(* IEC 61131-3 sources: codesys-elevator/codesys/src, 10 files *)

(* ---- E_Direction.st ---- *)
(* ==========================================================================
   E_Direction : かごの進行方向（Modbus の IR3 にそのまま載る）
   ========================================================================== *)
{attribute 'qualified_only'}   (* CODESYS 独自: E_Direction.Up の形でしか書けないようにする *)
TYPE E_Direction :
(
    Stop := 0,
    Up   := 1,
    Down := 2
) INT;
END_TYPE

(* ---- E_ElevCmd.st ---- *)
(* ==========================================================================
   E_ElevCmd : 画面から送られてくる指令の種類（Modbus の HR0 の値）
   ========================================================================== *)
{attribute 'qualified_only'}   (* CODESYS 独自: E_ElevCmd.CarCall の形でしか書けないようにする *)
TYPE E_ElevCmd :
(
    None      := 0,
    CarCall   := 1,   (* かご内の行き先ボタン（対象階 = HR1） *)
    HallCall  := 2,   (* 乗り場の呼びボタン（対象階 = HR1） *)
    DoorOpen  := 3,   (* 「開」ボタン *)
    DoorClose := 4    (* 「閉」ボタン *)
) INT;
END_TYPE

(* ---- E_ElevState.st ---- *)
(* ==========================================================================
   E_ElevState : エレベータの状態
   値は Modbus の IR0 にそのまま載り、画面（web/src/config.ts）と対応しているので、
   番号を変えないこと
   ========================================================================== *)
{attribute 'qualified_only'}   (* CODESYS 独自: E_ElevState.Idle の形でしか書けないようにする *)
TYPE E_ElevState :
(
    Idle        := 0,   (* 扉を閉めて停止中 *)
    DoorOpening := 1,   (* 扉を開けている途中 *)
    DoorOpen    := 2,   (* 扉が開いている（乗り降り中） *)
    DoorClosing := 3,   (* 扉を閉めている途中 *)
    Moving      := 4,   (* 移動中 *)
    Overload    := 5    (* 重量・人数オーバー。扉を開けたまま警報 *)
) INT;
END_TYPE

(* ---- GVL_ElevIO.st ---- *)
(* ==========================================================================
   GVL_ElevIO : Modbus TCP Slave の I/O マッピング先
   ・aElevToTS   → ModbusTCP Slave の「Input Registers」(%QW) にマッピング（20 個）
   ・aElevFromTS → ModbusTCP Slave の「Holding Registers」(%IW) にマッピング（10 個）
   各レジスタの意味は README.md のレジスタマップ表を参照
   ========================================================================== *)
{attribute 'qualified_only'}   (* CODESYS 独自: GVL_ElevIO.aElevToTS の形でしか書けないようにする *)
VAR_GLOBAL
    aElevToTS   : ARRAY[0..19] OF WORD;   (* PLC → TypeScript（FC04 で読まれる） *)
    aElevFromTS : ARRAY[0..9]  OF WORD;   (* TypeScript → PLC（FC16 で書かれる） *)
END_VAR

(* ---- GVL_ElevParam.st ---- *)
(* ==========================================================================
   GVL_ElevParam : エレベータの仕様（定数）
   画面側（web/src/config.ts）は IR11〜13 で受け取った値を使うので、
   ここを変えれば画面も追従する（FLOOR_COUNT は最大 16）
   ========================================================================== *)
{attribute 'qualified_only'}   (* CODESYS 独自: GVL_ElevParam.FLOOR_COUNT の形でしか書けないようにする *)
VAR_GLOBAL CONSTANT
    FLOOR_COUNT        : INT  := 5;       (* 階数 [階]。1F〜5F。呼びは WORD のビットで持つので最大 16 *)
    MAX_LOAD_KG        : INT  := 600;     (* 定格積載量 [kg] *)
    MAX_PERSONS        : INT  := 9;       (* 定員 [人] *)
    SPEED_FLOORS_PER_S : REAL := 0.5;     (* かごの速さ [階/s] *)
    DOOR_TRAVEL        : TIME := T#2S;    (* 扉が全閉から全開になるまでの時間 *)
    DOOR_DWELL         : TIME := T#5S;    (* 扉を開けておく時間（閉ボタンで短縮できる） *)
    POSITION_EPS       : REAL := 0.001;   (* 階に着いたかの判定の許容差 [階] *)
END_VAR

(* ---- FC_FloorBit.st ---- *)
(* ==========================================================================
   FC_FloorBit
   目的 : 階番号を、呼びを表す WORD のビットに変換する（bit0 = 1F）
   入力 : nFloor  階 [1..FLOOR_COUNT]
   戻り : 該当ビットだけ立った WORD。範囲外の階は 0（呼びとして扱わない）
   履歴 : 2026-10-19  初版
   ========================================================================== *)
FUNCTION FC_FloorBit : WORD
VAR_INPUT
    nFloor : INT;
END_VAR

IF nFloor >= 1 AND nFloor <= GVL_ElevParam.FLOOR_COUNT THEN
    FC_FloorBit := SHL(WORD#1, nFloor - 1);
ELSE
    FC_FloorBit := 0;   (* 画面から範囲外の階が来ても、存在しない階を呼ばない *)
END_IF

(* ---- FC_NextCallFloor.st ---- *)
(* ==========================================================================
   FC_NextCallFloor
   目的 : 進行方向の先にある、いちばん近い呼びの階を探す
          （エレベータの基本的な運転方式：今の方向の呼びを順に片付けてから折り返す）
   入力 : wCalls      呼び（かご内 OR 乗り場。bit0 = 1F）
          rPosition   かごの現在位置 [階]
          eDirection  探す方向
   戻り : 見つかった階 [1..FLOOR_COUNT]。無ければ 0
   履歴 : 2026-10-19  初版
   ========================================================================== *)
FUNCTION FC_NextCallFloor : INT
VAR_INPUT
    wCalls     : WORD;
    rPosition  : REAL;
    eDirection : E_Direction;
END_VAR
VAR
    nFloor : INT;
END_VAR

FC_NextCallFloor := 0;

CASE eDirection OF
    E_Direction.Up:
        (* 下から順に見て、今の位置以上で最初に見つかった呼び *)
        FOR nFloor := 1 TO GVL_ElevParam.FLOOR_COUNT DO
            IF (wCalls AND FC_FloorBit(nFloor)) <> 0
               AND INT_TO_REAL(nFloor) >= rPosition - GVL_ElevParam.POSITION_EPS THEN
                FC_NextCallFloor := nFloor;
                RETURN;
            END_IF
        END_FOR

    E_Direction.Down:
        (* 上から順に見て、今の位置以下で最初に見つかった呼び *)
        FOR nFloor := GVL_ElevParam.FLOOR_COUNT TO 1 BY -1 DO
            IF (wCalls AND FC_FloorBit(nFloor)) <> 0
               AND INT_TO_REAL(nFloor) <= rPosition + GVL_ElevParam.POSITION_EPS THEN
                FC_NextCallFloor := nFloor;
                RETURN;
            END_IF
        END_FOR

ELSE
    ;   (* 停止方向には「先」が無い *)
END_CASE

(* ---- FB_Door.st ---- *)
(* ==========================================================================
   FB_Door
   目的 : エレベータの扉の開閉の動きを模擬する
          （実機ならドア駆動装置への指令と、全開・全閉リミットスイッチの入力になる）
   入力 : bOpen    TRUE の間は開く方向、FALSE の間は閉じる方向へ動く
          tTravel  全閉から全開までの時間
          tDelta   前回呼んでからの経過時間
   出力 : nPositionPct  開き具合 [%]（0 = 全閉、100 = 全開）
          bIsOpen / bIsClosed  全開・全閉
   履歴 : 2026-10-19  初版
   ========================================================================== *)
FUNCTION_BLOCK FB_Door
VAR_INPUT
    bOpen   : BOOL;
    tTravel : TIME := T#2S;
    tDelta  : TIME;
END_VAR
VAR_OUTPUT
    nPositionPct : INT;
    bIsOpen      : BOOL;
    bIsClosed    : BOOL := TRUE;
END_VAR
VAR
    rPosition : REAL;   (* 0.0 = 全閉、1.0 = 全開 *)
    rStep     : REAL;
END_VAR

IF tTravel > T#0S THEN
    rStep := TIME_TO_REAL(tDelta) / TIME_TO_REAL(tTravel);
ELSE
    rStep := 1.0;       (* 時間 0 指定なら即座に動き切る *)
END_IF

IF bOpen THEN
    rPosition := MIN(1.0, rPosition + rStep);
ELSE
    rPosition := MAX(0.0, rPosition - rStep);
END_IF

nPositionPct := REAL_TO_INT(rPosition * 100.0);
bIsOpen      := nPositionPct >= 100;
bIsClosed    := nPositionPct <= 0;

(* ---- FB_Elevator.st ---- *)
(* ==========================================================================
   FB_Elevator
   目的 : エレベータ1台の制御（呼びの受け付け、運転方向の決定、扉、重量超過）
          グローバル変数には触らず、入出力だけでやり取りする（I/O は PRG_Elevator が担当）
   入力 : bCmdNew    新しい指令が来たサイクルだけ TRUE
          eCmd       指令の種類
          nCmdFloor  指令の対象階 [1..FLOOR_COUNT]
          nPersons   かごに乗っている人数 [人]
          nLoadKg    かごの積載重量 [kg]
          tDelta     前回呼んでからの経過時間
   出力 : eState, eDirection, rPosition [階], nFloor, nDoorPct [%],
          wCarCalls / wHallCalls（bit0 = 1F）, bOverload
   動き : ・呼ばれた階に向かい、着いたら扉を開ける
          ・扉は DOOR_DWELL だけ開けて閉じる（閉ボタンで短縮、開ボタンで延長）
          ・扉が開いている間に重量・人数が定格を超えたら Overload（扉を開けたまま警報）
          ・運転方向は「今の方向の呼びを片付けてから折り返す」
   履歴 : 2026-10-19  初版
   ========================================================================== *)
FUNCTION_BLOCK FB_Elevator
VAR_INPUT
    bCmdNew   : BOOL;
    eCmd      : E_ElevCmd;
    nCmdFloor : INT;
    nPersons  : INT;
    nLoadKg   : INT;
    tDelta    : TIME;
END_VAR
VAR_OUTPUT
    eState     : E_ElevState := E_ElevState.Idle;
    eDirection : E_Direction := E_Direction.Stop;
    rPosition  : REAL := 1.0;   (* 1.0 = 1F *)
    nFloor     : INT := 1;      (* いちばん近い階 *)
    nDoorPct   : INT;
    wCarCalls  : WORD;
    wHallCalls : WORD;
    bOverload  : BOOL;
END_VAR
VAR
    fbDoor           : FB_Door;
    tonDwell         : TON;
    eTravelDirection : E_Direction := E_Direction.Up;   (* 走行中の方向。停止中は次に優先して探す方向 *)
    wCarCallIn       : WORD;    (* このサイクルに押されたボタン *)
    wHallCallIn      : WORD;
    wAllCalls        : WORD;
    wAnswered        : WORD;    (* このサイクルに応答した（消す）呼び *)
    bOpenRequest     : BOOL;
    bCloseRequest    : BOOL;
    nTarget          : INT;
    rStep            : REAL;
    rNext            : REAL;
END_VAR

(* ---- 指令の受け付け（このサイクルの分だけ） ---- *)
wCarCallIn    := SEL(bCmdNew AND eCmd = E_ElevCmd.CarCall,  WORD#0, FC_FloorBit(nCmdFloor));
wHallCallIn   := SEL(bCmdNew AND eCmd = E_ElevCmd.HallCall, WORD#0, FC_FloorBit(nCmdFloor));
bOpenRequest  := bCmdNew AND eCmd = E_ElevCmd.DoorOpen;
bCloseRequest := bCmdNew AND eCmd = E_ElevCmd.DoorClose;

wAllCalls := wCarCalls OR wHallCalls OR wCarCallIn OR wHallCallIn;
bOverload := nLoadKg > GVL_ElevParam.MAX_LOAD_KG OR nPersons > GVL_ElevParam.MAX_PERSONS;
wAnswered := 0;

(* 扉を開けておく時間。DoorOpen 以外では IN が FALSE になり、自動でリセットされる *)
tonDwell(IN := eState = E_ElevState.DoorOpen, PT := GVL_ElevParam.DOOR_DWELL);

(* ---- 状態遷移 ---- *)
CASE eState OF
    E_ElevState.Idle:
        IF bOpenRequest OR (wAllCalls AND FC_FloorBit(nFloor)) <> 0 THEN
            eState := E_ElevState.DoorOpening;              (* 今いる階で呼ばれた *)
        ELSIF FC_NextCallFloor(wAllCalls, rPosition, eTravelDirection) <> 0 THEN
            eState := E_ElevState.Moving;                    (* 前と同じ方向に呼びがある *)
        ELSIF wAllCalls <> 0 THEN
            (* 同じ方向に呼びが無い → 折り返す *)
            IF eTravelDirection = E_Direction.Up THEN
                eTravelDirection := E_Direction.Down;
            ELSE
                eTravelDirection := E_Direction.Up;
            END_IF
            eState := E_ElevState.Moving;
        END_IF

    E_ElevState.DoorOpening:
        wAnswered := FC_FloorBit(nFloor);                    (* この階の呼びに応答した *)
        IF fbDoor.bIsOpen THEN
            eState := E_ElevState.DoorOpen;
        END_IF

    E_ElevState.DoorOpen:
        wAnswered := FC_FloorBit(nFloor);
        IF bOverload THEN
            eState := E_ElevState.Overload;
        ELSIF bOpenRequest THEN
            eState := E_ElevState.DoorOpening;   (* 開ボタン: 一度抜けることで待ち時間をやり直す *)
        ELSIF tonDwell.Q OR bCloseRequest THEN
            eState := E_ElevState.DoorClosing;
        END_IF

    E_ElevState.Overload:
        wAnswered := FC_FloorBit(nFloor);
        IF NOT bOverload THEN
            eState := E_ElevState.DoorOpen;      (* 降りて定格内に戻ったら、待ち時間から再開 *)
        END_IF

    E_ElevState.DoorClosing:
        (* 閉まりかけでも、開ボタン・この階の呼び・駆け込みによる超過があれば開け直す *)
        IF bOpenRequest OR bOverload OR (wAllCalls AND FC_FloorBit(nFloor)) <> 0 THEN
            eState := E_ElevState.DoorOpening;
        ELSIF fbDoor.bIsClosed THEN
            eState := E_ElevState.Idle;          (* 次の行き先は Idle で決める *)
        END_IF

    E_ElevState.Moving:
        nTarget := FC_NextCallFloor(wAllCalls, rPosition, eTravelDirection);
        IF nTarget = 0 THEN
            (* 呼びは着くまで消えないので通常は起きない。念のため次の階で止める *)
            IF eTravelDirection = E_Direction.Up THEN
                nTarget := LIMIT(1, DINT_TO_INT(TRUNC(rPosition)) + 1, GVL_ElevParam.FLOOR_COUNT);
            ELSE
                nTarget := LIMIT(1, DINT_TO_INT(TRUNC(rPosition)), GVL_ElevParam.FLOOR_COUNT);
            END_IF
        END_IF

        rStep := GVL_ElevParam.SPEED_FLOORS_PER_S * TIME_TO_REAL(tDelta) / 1000.0;
        IF eTravelDirection = E_Direction.Up THEN
            rNext := rPosition + rStep;
            IF rNext >= INT_TO_REAL(nTarget) THEN
                rNext  := INT_TO_REAL(nTarget);   (* 行き過ぎないよう階にぴったり合わせる *)
                eState := E_ElevState.DoorOpening;
            END_IF
        ELSE
            rNext := rPosition - rStep;
            IF rNext <= INT_TO_REAL(nTarget) THEN
                rNext  := INT_TO_REAL(nTarget);
                eState := E_ElevState.DoorOpening;
            END_IF
        END_IF
        rPosition := rNext;

ELSE
    (* 列挙外の値はメモリ破壊などの異常。走行を止め、扉を閉めた停止状態に戻す *)
    eState := E_ElevState.Idle;
END_CASE

(* ---- 出力（ここでまとめて決める） ---- *)
fbDoor(bOpen := eState = E_ElevState.DoorOpening
             OR eState = E_ElevState.DoorOpen
             OR eState = E_ElevState.Overload,
       tTravel := GVL_ElevParam.DOOR_TRAVEL,
       tDelta := tDelta);
nDoorPct := fbDoor.nPositionPct;

wCarCalls  := (wCarCalls  OR wCarCallIn)  AND NOT wAnswered;
wHallCalls := (wHallCalls OR wHallCallIn) AND NOT wAnswered;

nFloor := LIMIT(1, REAL_TO_INT(rPosition), GVL_ElevParam.FLOOR_COUNT);

IF eState = E_ElevState.Moving THEN
    eDirection := eTravelDirection;
ELSE
    eDirection := E_Direction.Stop;
END_IF

(* ---- PRG_Elevator.st ---- *)
(* ==========================================================================
   PRG_Elevator
   目的 : Modbus のレジスタ（GVL_ElevIO）と FB_Elevator の橋渡し
          グローバル変数を触るのはこのプログラムだけにする
   入力 : GVL_ElevIO.aElevFromTS[0..4]  指令（種類・階・通し番号）、人数、重量
   出力 : GVL_ElevIO.aElevToTS[0..14]   状態、位置、扉、呼び、警報、定格値など
          （各レジスタの意味は README.md のレジスタマップ表を参照）
   指令 : 画面は「種類・階・通し番号」を1回の書き込み（FC16）で送る。
          通し番号が前回と変わったサイクルだけ、新しい指令として扱う
          （同じ階のボタンを2回押しても取りこぼさないため）
   使い方 : MainTask から毎サイクル呼ぶ
   履歴 : 2026-10-19  初版
   ========================================================================== *)
PROGRAM PRG_Elevator
VAR CONSTANT
    MAX_DELTA      : TIME := T#100MS;   (* 停止明けなどで経過時間が飛んだときの上限 *)
    POSITION_SCALE : REAL := 100.0;     (* 位置 [階] を INT に詰める倍率（1.00F → 100） *)
    MAX_INPUT      : INT  := 9999;      (* 人数・重量として受け付ける上限 *)
END_VAR
VAR
    fbElevator  : FB_Elevator;
    eCmdIn      : E_ElevCmd;
    nLastSeq    : WORD;
    bFirstCycle : BOOL := TRUE;
    tNow        : TIME;
    tLast       : TIME;
    tDelta      : TIME;
    wHeartbeat  : WORD;
END_VAR

(* ---- 経過時間 ---- *)
tNow := TIME();                        (* 起動からの経過時間 *)
IF bFirstCycle THEN
    tDelta   := T#0S;
    nLastSeq := GVL_ElevIO.aElevFromTS[2];   (* 起動前に残っていた指令は実行しない *)
ELSIF tNow - tLast > MAX_DELTA THEN
    tDelta := MAX_DELTA;
ELSE
    tDelta := tNow - tLast;
END_IF
tLast := tNow;
bFirstCycle := FALSE;

(* ---- 指令の種類（範囲外の値は None にして無視する） ---- *)
CASE WORD_TO_INT(GVL_ElevIO.aElevFromTS[0]) OF
    1: eCmdIn := E_ElevCmd.CarCall;
    2: eCmdIn := E_ElevCmd.HallCall;
    3: eCmdIn := E_ElevCmd.DoorOpen;
    4: eCmdIn := E_ElevCmd.DoorClose;
ELSE
    eCmdIn := E_ElevCmd.None;
END_CASE

(* ---- 制御本体 ---- *)
fbElevator(
    bCmdNew   := GVL_ElevIO.aElevFromTS[2] <> nLastSeq,
    eCmd      := eCmdIn,
    nCmdFloor := WORD_TO_INT(GVL_ElevIO.aElevFromTS[1]),
    nPersons  := LIMIT(0, WORD_TO_INT(GVL_ElevIO.aElevFromTS[3]), MAX_INPUT),
    nLoadKg   := LIMIT(0, WORD_TO_INT(GVL_ElevIO.aElevFromTS[4]), MAX_INPUT),
    tDelta    := tDelta);
nLastSeq := GVL_ElevIO.aElevFromTS[2];

(* ---- 画面へ出す値 ---- *)
wHeartbeat := wHeartbeat + 1;   (* 通信の生存確認用。WORD なので 65535 の次は 0 に戻ってよい *)

GVL_ElevIO.aElevToTS[0]  := INT_TO_WORD(fbElevator.eState);
GVL_ElevIO.aElevToTS[1]  := INT_TO_WORD(REAL_TO_INT(fbElevator.rPosition * POSITION_SCALE));
GVL_ElevIO.aElevToTS[2]  := INT_TO_WORD(fbElevator.nFloor);
GVL_ElevIO.aElevToTS[3]  := INT_TO_WORD(fbElevator.eDirection);
GVL_ElevIO.aElevToTS[4]  := INT_TO_WORD(fbElevator.nDoorPct);
GVL_ElevIO.aElevToTS[5]  := fbElevator.wCarCalls;
GVL_ElevIO.aElevToTS[6]  := fbElevator.wHallCalls;
GVL_ElevIO.aElevToTS[7]  := INT_TO_WORD(LIMIT(0, WORD_TO_INT(GVL_ElevIO.aElevFromTS[3]), MAX_INPUT));
GVL_ElevIO.aElevToTS[8]  := INT_TO_WORD(LIMIT(0, WORD_TO_INT(GVL_ElevIO.aElevFromTS[4]), MAX_INPUT));
(* 状態フラグ: bit0 超過 / bit1 警報中 / bit2 扉全開 / bit3 扉全閉 / bit4 移動中 *)
GVL_ElevIO.aElevToTS[9]  := BOOL_TO_WORD(fbElevator.bOverload)
                         OR SHL(BOOL_TO_WORD(fbElevator.eState = E_ElevState.Overload), 1)
                         OR SHL(BOOL_TO_WORD(fbElevator.nDoorPct >= 100), 2)
                         OR SHL(BOOL_TO_WORD(fbElevator.nDoorPct <= 0), 3)
                         OR SHL(BOOL_TO_WORD(fbElevator.eState = E_ElevState.Moving), 4);
GVL_ElevIO.aElevToTS[10] := nLastSeq;   (* 処理済みの通し番号（画面が受け付けを確認する） *)
GVL_ElevIO.aElevToTS[11] := INT_TO_WORD(GVL_ElevParam.MAX_LOAD_KG);
GVL_ElevIO.aElevToTS[12] := INT_TO_WORD(GVL_ElevParam.MAX_PERSONS);
GVL_ElevIO.aElevToTS[13] := INT_TO_WORD(GVL_ElevParam.FLOOR_COUNT);
GVL_ElevIO.aElevToTS[14] := wHeartbeat;
